VAR_GLOBAL

	eLightTowerState: E_LightTowerState;
	eBuzzerMode: E_BuzzerMode;
	bBuzzerMute: BOOL;

	bPauseMachine: BOOL;
	bResumeMachine: BOOL;
	bResetAllCycles: BOOL;
	
	PauseAll: BOOL;
	PauseAllDelayed: BOOL;
	ResumeAll: BOOL;	

	iActErrors							: INT;
	iActMessages						: INT;
	iActWarning							: INT;

	fbMode	: ARRAY[0..E_ModeZone.eLast] OF FB_ModeSelect;
	stMode	: ARRAY[0..E_ModeZone.eLast] OF ST_Mode;
	stOper	: ARRAY[0..E_ModeZone.eLast] OF ST_OperationButtons;
	
	fbLightTower: ARRAY[0..E_SkidZone.eLast] OF FB_LightTower;
	fbLightTower_Control: ARRAY[0..E_SkidZone.eLast] OF FB_LightTower_Control;



	//Operational Modes	
	stModeMain: ST_Mode;
	
	// Operational Buttons
	stOpMain				:ST_OperationButtons;
	stOpNonPause			:ST_OperationButtons;	

END_VAR

(* stored: Version 1.1.0.1, ProductVersion 3.1.4024.15
   GVL GVL_OperMode: Id {db8bfe85-e73f-4c80-9836-be8123e81b8e} *)
